//Get read/write access to content
//Get_P returns a pointer to the Dummy instance
METHOD PROTECTED _Get_P : POINTER TO FB_processStep_Flow

VAR_INPUT
	NumberOfObject	: UDINT;
	Response				: REFERENCE TO KOSTAL_TC3_Core_functionResponse.FB_functionResponse;
END_VAR

VAR
	_response: KOSTAL_TC3_Core_functionResponse.FB_functionResponse;
END_VAR

_response.clear();

IF (NumberOfObject = 0) 
OR (NumberOfObject > _ListOfObject.nObjects)
OR (_ListOfObject.pObjects = 0)
THEN

	_Dummy.Clear();

	_Get_P:= ADR(_Dummy);

	_response.status:= 'return Dummy because NumberOfPosition is out of range';

ELSE

	_response.success:= TRUE;
	
	_Get_P:= _ListOfObject.pObjects[NumberOfObject - 1];

END_IF

IF __ISVALIDREF(Response) THEN	Response.CopyFrom(_response);	END_IF
END_METHOD

//Overwrites the method in the base class with the real contents of the ListOf class.
METHOD PROTECTED  _New : PVOID

VAR
	_pNew: POINTER TO FB_processStep_Flow;
END_VAR

_pNew:= __NEW(FB_processStep_Flow);

_New:= _pNew;
END_METHOD

//Add a new instance of FB_Dut and copy content from [IN] to the new instance
METHOD PUBLIC Add_DUT : BOOL
VAR_INPUT
	IN				: I_processStep_Flow;
	Response	: REFERENCE TO KOSTAL_TC3_Core_functionResponse.FB_functionResponse;
END_VAR

VAR
	pDUT: POINTER TO FB_processStep_Flow;
	_response: KOSTAL_TC3_Core_functionResponse.FB_functionResponse;
END_VAR
_response.clear();

//create a new empty object 
IF NOT _AddObject() THEN
	_response.status:= ('_AddObject failed');
	IF __ISVALIDREF(Response) THEN	Response.CopyFrom(_response);	END_IF
	RETURN;	
END_IF

//Return, if no  [IN] object is available
IF IN = 0 THEN 
	_response.status:= ('IN Parameter not defined');
	IF __ISVALIDREF(Response) THEN	Response.CopyFrom(_response);	END_IF
	RETURN;	
END_IF

//otherwise fill [IN] object content to new virtual instance
pDUT:= _Get_P(_ListOfObject.nObjects, _response);

IF NOT _response.success THEN 
	IF __ISVALIDREF(Response) THEN	Response.CopyFrom(_response);	END_IF
	RETURN;	
END_IF

IF pDUT = 0 THEN 
	_response.status:= ('no Pointer get from list');
	IF __ISVALIDREF(Response) THEN	Response.CopyFrom(_response);	END_IF
	RETURN;	
END_IF

pDut^.CopyFrom(IN);

_response.success:= TRUE;
IF __ISVALIDREF(Response) THEN	Response.CopyFrom(_response);	END_IF

Add_DUT:= TRUE;
END_METHOD

METHOD PUBLIC CopyFrom
VAR_INPUT
	IN	: I_ListOf_processStep_Flow;
END_VAR

VAR
	_udi: UDINT;
END_VAR

IF IN = 0 THEN RETURN;	END_IF

Clear();

FOR _udi:= 1 TO IN.NumberOfObjects DO
	Add_DUT(IN.Get_I(_udi, 0), 0);
END_FOR
END_METHOD

METHOD PUBLIC CopyTo
VAR_INPUT
	IN	: I_ListOf_processStep_Flow_CopyFrom;
END_VAR

IF IN = 0 THEN RETURN;	END_IF

IN.CopyFrom(THIS^);
END_METHOD

METHOD PUBLIC Delete_DUT : BOOL
VAR_INPUT
	Number	: UDINT;	//Number of DUT in List
END_VAR

VAR
	_Set: FB_ListOf_processStep_Flow;
	_udi: UDINT;
END_VAR

//Range control
IF Number = 0 							THEN RETURN;	END_IF
IF Number > NumberOfObjects	THEN RETURN;	END_IF

//Intermediate storage - prepare
_Set.Clear();

//catch all elements without the Number defiend
FOR _udi:= 1 TO NumberOfObjects DO
	IF _udi <> Number THEN
		_Set.Add_DUT(THIS^.Get_I(_udi, 0), 0);
	END_IF
END_FOR

//Delete own content
Clear();

//Add the remaining elements of the own class. 
FOR _udi:= 1 TO _Set.NumberOfObjects DO
		THIS^.Add_DUT(_Set.Get_I(_udi, 0), 0);
END_FOR

//Intermediate storage - clean Router storage
_Set.Clear();

Delete_DUT:= TRUE;
END_METHOD

//Get readonly access to content 
METHOD Get_I : I_processStep_Flow

VAR_INPUT
	NumberOfObject	: UDINT;
	Response				: REFERENCE TO KOSTAL_TC3_Core_functionResponse.FB_functionResponse;
END_VAR

VAR
	_response: KOSTAL_TC3_Core_functionResponse.FB_functionResponse;
END_VAR

_response.clear();

Get_I:= _Get_P(NumberOfObject, _response)^;

IF __ISVALIDREF(Response) THEN	Response.CopyFrom(_response);	END_IF
END_METHOD

//Get full access to content 
METHOD Get_IOwner : I_processStep_Flow_Owner

VAR_INPUT
	NumberOfObject	: UDINT;
	Response				: REFERENCE TO KOSTAL_TC3_Core_functionResponse.FB_functionResponse;
END_VAR

VAR
	_response: KOSTAL_TC3_Core_functionResponse.FB_functionResponse;
END_VAR

_response.clear();

Get_IOwner:= _Get_P(NumberOfObject, _response)^;

IF __ISVALIDREF(Response) THEN	Response.CopyFrom(_response);	END_IF
END_METHOD

END_FUNCTION_BLOCK

// Step/DUT/processStep_Flow/ListOf/I_ListOf_processStep_Flow
INTERFACE I_ListOf_processStep_Flow EXTENDS KOSTAL_TC3_Components_ListOf_Objects.I_Base

METHOD PUBLIC CopyTo
VAR_INPUT
	IN	: I_ListOf_processStep_Flow_CopyFrom;
END_VAR
END_METHOD

METHOD Get_I : I_processStep_Flow

VAR_INPUT
	NumberOfObject	: UDINT;
	Response				: REFERENCE TO KOSTAL_TC3_Core_functionResponse.FB_functionResponse;
END_VAR
END_METHOD

END_INTERFACE

// Step/DUT/processStep_Flow/ListOf/I_ListOf_processStep_Flow_CopyFrom
INTERFACE I_ListOf_processStep_Flow_CopyFrom EXTENDS KOSTAL_TC3_Core_System.I_Interface

METHOD PUBLIC CopyFrom
VAR_INPUT
	IN	: I_ListOf_processStep_Flow;
END_VAR
END_METHOD

END_INTERFACE

// Step/DUT/processStep_Flow/I_processStep_Flow
INTERFACE I_processStep_Flow EXTENDS I_processStep

METHOD PUBLIC isCalledExternally : BOOL
VAR_INPUT
END_VAR
END_METHOD

METHOD PUBLIC NotFound : BOOL
VAR_INPUT
END_VAR
END_METHOD

END_INTERFACE

// Step/DUT/processStep_Flow/ListOf/I_ListOf_processStep_Flow_Owner
INTERFACE I_ListOf_processStep_Flow_Owner EXTENDS KOSTAL_TC3_Components_ListOf_Objects.I_Base_Owner

//Add a new instance of FB_Dut and copy content from [IN] to the new instance
METHOD PUBLIC Add_DUT : BOOL
VAR_INPUT
	IN				: I_processStep_Flow;
	Response	: REFERENCE TO KOSTAL_TC3_Core_functionResponse.FB_functionResponse;
END_VAR
END_METHOD

METHOD PUBLIC CopyFrom
VAR_INPUT
	IN	: I_ListOf_processStep_Flow;
END_VAR
END_METHOD

METHOD PUBLIC CopyTo
VAR_INPUT
	IN	: I_ListOf_processStep_Flow_CopyFrom;
END_VAR
END_METHOD

METHOD PUBLIC Delete_DUT : BOOL
VAR_INPUT
	Number	: UDINT;	//Number of DUT in List
END_VAR
END_METHOD

//Get readonly access to content 
METHOD Get_I : I_processStep_Flow

VAR_INPUT
	NumberOfObject	: UDINT;
	Response				: REFERENCE TO KOSTAL_TC3_Core_functionResponse.FB_functionResponse;
END_VAR
END_METHOD

//Get full access to content 
METHOD Get_IOwner : I_processStep_Flow_Owner

VAR_INPUT
	NumberOfObject	: UDINT;
	Response				: REFERENCE TO KOSTAL_TC3_Core_functionResponse.FB_functionResponse;
END_VAR
END_METHOD

END_INTERFACE

// Step/DUT/processStep_Flow/I_processStep_Flow_Owner
INTERFACE I_processStep_Flow_Owner EXTENDS I_processStep_Owner

METHOD PUBLIC clear
END_METHOD

(*
Description
===========
| Apply changes in step sequence
| Call before or after the step sequence (see usage sample)
*)
METHOD PUBLIC Header
VAR_INPUT
END_VAR
END_METHOD

(*
Description
===========
| Reset step sequence to 0
*)
METHOD PUBLIC init
END_METHOD

(*
| Description
| ============
| Returns TRUE if step.active is equal stepNumber 
*)

METHOD PUBLIC isActive : BOOL
VAR_INPUT
	stepNumber	: INT;
END_VAR
END_METHOD

METHOD PUBLIC isCalledExternally : BOOL
VAR_INPUT
END_VAR
END_METHOD

METHOD PUBLIC NotFound : BOOL
VAR_INPUT
END_VAR
END_METHOD

END_INTERFACE

// Step/DUT/processStep_Flow/FB_processStep_Flow
(*

:Author: Frank Dümpelmann <f.duempelmann@kostal.com>
:Date: 2019-03-29

Function
========
| Extends FB_processStep

Methods and Properties
======================
| See bottom of this document for a detailed description of each method or property
*)

{attribute 'enable_dynamic_creation'}
FUNCTION_BLOCK PUBLIC FB_processStep_Flow EXTENDS FB_processStep IMPLEMENTS I_processStep_Flow, I_processStep_Flow_Owner

VAR
	_Found	: BOOL;
END_VAR

METHOD PUBLIC clear

_Found:= FALSE;

SUPER^.clear();
END_METHOD

(*
Description
===========
| Apply changes in step sequence
| Call before or after the step sequence (see usage sample)
*)
METHOD PUBLIC Header
VAR_INPUT
END_VAR

_Found:= FALSE;
END_METHOD

(*
Description
===========
| Reset step sequence to 0
*)
METHOD PUBLIC init

_Found:= FALSE;

SUPER^.init();
END_METHOD

(*
| Description
| ============
| Returns TRUE if step.active is equal stepNumber 
*)

METHOD PUBLIC isActive : BOOL
VAR_INPUT
	stepNumber	: INT;
END_VAR
 
isActive:= _request = stepNumber;

IF NOT isActive THEN RETURN;	END_IF

_Found:= TRUE;

SUPER^.Header();
END_METHOD

METHOD PUBLIC isCalledExternally : BOOL
VAR_INPUT
END_VAR

isCalledExternally:= _actual <> _request;
END_METHOD

METHOD PUBLIC NotFound : BOOL
VAR_INPUT
END_VAR

NotFound:= NOT _Found;
END_METHOD

END_FUNCTION_BLOCK

// Step/POE/ListOf/FB_ListOf_ProcessStep_Control
FUNCTION_BLOCK FB_ListOf_ProcessStep_Control  EXTENDS KOSTAL_TC3_Components_ListOf_Objects.FB_Base IMPLEMENTS I_ListOf_ProcessStep_Control, I_ListOf_ProcessStep_Control_CopyFrom, I_ListOf_ProcessStep_Control_Owner

VAR
	_Dummy	: FB_ProcessStep_Control;
END_VAR

//Overwrites the method in the base class with the real contents of the ListOf class.
METHOD PROTECTED  _deletePayLoad
VAR_INPUT
	pPayload	:	PVOID; 
END_VAR

VAR
	_p	: POINTER TO FB_ProcessStep_Control;
END_VAR

IF pPayload = 0  THEN	RETURN;	END_IF

_p:= pPayload;

__DELETE(_p);
END_METHOD

//Get read/write access to content
//Get_P returns a pointer to the Dummy instance
METHOD PROTECTED _Get_P : POINTER TO FB_ProcessStep_Control

VAR_INPUT
	NumberOfObject	: UDINT;
	Response				: REFERENCE TO KOSTAL_TC3_Core_functionResponse.FB_functionResponse;
END_VAR

VAR
	_response: KOSTAL_TC3_Core_functionResponse.FB_functionResponse;
END_VAR

_response.clear();

IF (NumberOfObject = 0) 
OR (NumberOfObject > _ListOfObject.nObjects)
OR (_ListOfObject.pObjects = 0)
THEN

	//_Dummy.Clear(); No clean-up method 

	_Get_P:= ADR(_Dummy);

	_response.status:= 'return Dummy because NumberOfPosition is out of range';

ELSE

	_response.success:= TRUE;
	
	_Get_P:= _ListOfObject.pObjects[NumberOfObject - 1];

END_IF

IF __ISVALIDREF(Response) THEN	Response.CopyFrom(_response);	END_IF
END_METHOD

//Overwrites the method in the base class with the real contents of the ListOf class.
METHOD PROTECTED  _New : PVOID

VAR
	_pNew: POINTER TO FB_ProcessStep_Control;
END_VAR

_pNew:= __NEW(FB_ProcessStep_Control);

_New:= _pNew;
END_METHOD

//Add a new instance of FB_Dut and copy content from [IN] to the new instance
METHOD PUBLIC Add_DUT : BOOL
VAR_INPUT
	IN				: I_ProcessStep_Control;
	Response	: REFERENCE TO KOSTAL_TC3_Core_functionResponse.FB_functionResponse;
END_VAR

VAR
	pDUT: POINTER TO FB_ProcessStep_Control;
	_response: KOSTAL_TC3_Core_functionResponse.FB_functionResponse;
END_VAR
_response.clear();

//create a new empty object 
IF NOT _AddObject() THEN
	_response.status:= ('_AddObject failed');
	IF __ISVALIDREF(Response) THEN	Response.CopyFrom(_response);	END_IF
	RETURN;	
END_IF

//Return, if no  [IN] object is available
IF IN = 0 THEN 
	_response.status:= ('IN Parameter not defined');
	IF __ISVALIDREF(Response) THEN	Response.CopyFrom(_response);	END_IF
	RETURN;	
END_IF

//otherwise fill [IN] object content to new virtual instance
pDUT:= _Get_P(_ListOfObject.nObjects, _response);

IF NOT _response.success THEN 
	IF __ISVALIDREF(Response) THEN	Response.CopyFrom(_response);	END_IF
	RETURN;	
END_IF

IF pDUT = 0 THEN 
	_response.status:= ('no Pointer get from list');
	IF __ISVALIDREF(Response) THEN	Response.CopyFrom(_response);	END_IF
	RETURN;	
END_IF

pDut^.CopyFrom(IN);

_response.success:= TRUE;
IF __ISVALIDREF(Response) THEN	Response.CopyFrom(_response);	END_IF

Add_DUT:= TRUE;
END_METHOD

METHOD PUBLIC CopyFrom
VAR_INPUT
	IN	: I_ListOf_ProcessStep_Control;
END_VAR

VAR
	_udi: UDINT;
END_VAR

IF IN = 0 THEN RETURN;	END_IF

Clear();

FOR _udi:= 1 TO IN.NumberOfObjects DO
	Add_DUT(IN.Get_I(_udi, 0), 0);
END_FOR
END_METHOD

METHOD PUBLIC CopyTo
VAR_INPUT
	IN	: I_ListOf_ProcessStep_Control_CopyFrom;
END_VAR

IF IN = 0 THEN RETURN;	END_IF

IN.CopyFrom(THIS^);
END_METHOD

METHOD PUBLIC Delete_DUT : BOOL
VAR_INPUT
	Number	: UDINT;	//Number of DUT in List
END_VAR

VAR
	_Set: FB_ListOf_ProcessStep_Control;
	_udi: UDINT;
END_VAR

//Range control
IF Number = 0 							THEN RETURN;	END_IF
IF Number > NumberOfObjects	THEN RETURN;	END_IF

//Intermediate storage - prepare
_Set.Clear();

//catch all elements without the Number defiend
FOR _udi:= 1 TO NumberOfObjects DO
	IF _udi <> Number THEN
		_Set.Add_DUT(THIS^.Get_I(_udi, 0), 0);
	END_IF
END_FOR

//Delete own content
Clear();

//Add the remaining elements of the own class. 
FOR _udi:= 1 TO _Set.NumberOfObjects DO
		THIS^.Add_DUT(_Set.Get_I(_udi, 0), 0);
END_FOR

//Intermediate storage - clean Router storage
_Set.Clear();

Delete_DUT:= TRUE;
END_METHOD

//Get readonly access to content 
METHOD Get_I : I_ProcessStep_Control

VAR_INPUT
	NumberOfObject	: UDINT;
	Response				: REFERENCE TO KOSTAL_TC3_Core_functionResponse.FB_functionResponse;
END_VAR

VAR
	_response: KOSTAL_TC3_Core_functionResponse.FB_functionResponse;
END_VAR

_response.clear();

Get_I:= _Get_P(NumberOfObject, _response)^;

IF __ISVALIDREF(Response) THEN	Response.CopyFrom(_response);	END_IF
END_METHOD

//Get full access to content 
METHOD Get_IOwner : I_ProcessStep_Control_Owner

VAR_INPUT
	NumberOfObject	: UDINT;
	Response				: REFERENCE TO KOSTAL_TC3_Core_functionResponse.FB_functionResponse;
END_VAR

VAR
	_response: KOSTAL_TC3_Core_functionResponse.FB_functionResponse;
END_VAR

_response.clear();

Get_IOwner:= _Get_P(NumberOfObject, _response)^;

IF __ISVALIDREF(Response) THEN	Response.CopyFrom(_response);	END_IF
END_METHOD

END_FUNCTION_BLOCK

// Step/POE/ListOf/I_ListOf_ProcessStep_Control
INTERFACE I_ListOf_ProcessStep_Control EXTENDS KOSTAL_TC3_Components_ListOf_Objects.I_Base

METHOD PUBLIC CopyTo
VAR_INPUT
	IN	: I_ListOf_ProcessStep_Control_CopyFrom;
END_VAR
END_METHOD

METHOD Get_I : I_ProcessStep_Control

VAR_INPUT
	NumberOfObject	: UDINT;
	Response				: REFERENCE TO KOSTAL_TC3_Core_functionResponse.FB_functionResponse;
END_VAR
END_METHOD

END_INTERFACE

// Step/POE/ListOf/I_ListOf_ProcessStep_Control_CopyFrom
INTERFACE I_ListOf_ProcessStep_Control_CopyFrom EXTENDS KOSTAL_TC3_Core_System.I_Interface

METHOD PUBLIC CopyFrom
VAR_INPUT
	IN	: I_ListOf_ProcessStep_Control;
END_VAR
END_METHOD

END_INTERFACE

// Step/POE/ListOf/I_ListOf_ProcessStep_Control_Owner
INTERFACE I_ListOf_ProcessStep_Control_Owner EXTENDS KOSTAL_TC3_Components_ListOf_Objects.I_Base_Owner

//Add a new instance of FB_Dut and copy content from [IN] to the new instance
METHOD PUBLIC Add_DUT : BOOL
VAR_INPUT
	IN				: I_ProcessStep_Control;
	Response	: REFERENCE TO KOSTAL_TC3_Core_functionResponse.FB_functionResponse;
END_VAR
END_METHOD

METHOD PUBLIC CopyFrom
VAR_INPUT
	IN	: I_ListOf_ProcessStep_Control;
END_VAR
END_METHOD

METHOD PUBLIC CopyTo
VAR_INPUT
	IN	: I_ListOf_ProcessStep_Control_CopyFrom;
END_VAR
END_METHOD

METHOD PUBLIC Delete_DUT : BOOL
VAR_INPUT
	Number	: UDINT;	//Number of DUT in List
END_VAR
END_METHOD

//Get readonly access to content 
METHOD Get_I : I_ProcessStep_Control

VAR_INPUT
	NumberOfObject	: UDINT;
	Response				: REFERENCE TO KOSTAL_TC3_Core_functionResponse.FB_functionResponse;
END_VAR
END_METHOD

//Get full access to content 
METHOD Get_IOwner : I_ProcessStep_Control_Owner

VAR_INPUT
	NumberOfObject	: UDINT;
	Response				: REFERENCE TO KOSTAL_TC3_Core_functionResponse.FB_functionResponse;
END_VAR
END_METHOD

END_INTERFACE
